(* IEC 61131-3 sources: moulding-cell-robot-interlock/plc/test/st, 1 file *)

(* ---- tb_bench.st ---- *)
(*
  TB_BENCH: self-checking test bench for the function block CELL_PLC.
  Generated by scripts/make_testbench.py from the cell model (cell/bench.py). Do not edit.

  One call is one scan of the block under test. For every scan of every case the bench applies the
  recorded input image (machine model and TP program of the repository, one PLC scan per step),
  calls its own instance of CELL_PLC and compares all outputs, the state and the fault code with
  the recorded values. A case fails at its first difference. Every case starts with a fresh instance.
  Cases: 7. Scans: 1616. Table rows (equal consecutive scans are merged): 332.
  Input bits of rowIn, from bit 0: iZA6_MouldClosed, iZA7_MouldOpenPosition, iZB2_EnableOperation, iZB3_EjectorBack, iZB4_EjectorForward, iSafetyOk, rbReqClose, rbReqEjFwd, rbReqEjBack, rbAtCut, rbPlaced, rbFault, rbAtWait, rbAreaFree, iCutClosed, iCutOpen, iNestFree, iGateClosedLocked, btnGateReq, btnReset.
  Output bits of rowExp, from bit 0: qA6_EnableMouldClosure, qB3_EnableEjectorBack, qB4_EnableEjectorForward, qB2_NoOperationWithImm, qRbImmAuto, qRbMouldOpen, qRbMouldClosed, qRbEjFwd, qRbEjBack, qRbCutDone, qRbPlaceFree, qRbCycleEnable, qRbPlaceAck, qCutClose, qConvIndex, qGateUnlock.
  rowSt = state + 16 * faultCode.
*)

FUNCTION_BLOCK TB_BENCH
VAR_INPUT
  enable : BOOL;
END_VAR
VAR_OUTPUT
  Done : BOOL;
  CasesTotal : INT;
  CasesRun : INT;
  CasesPassed : INT;
  CasesFailed : INT;
  FirstFailedCase : INT;
  FirstFailedCheck : INT;      (* scan number inside the failed case, from 1 *)
  CasePassBits : DWORD;        (* bit 0 = case 1 *)
END_VAR
VAR
  dut1 : CELL_PLC;
  dut2 : CELL_PLC;
  dut3 : CELL_PLC;
  dut4 : CELL_PLC;
  dut5 : CELL_PLC;
  dut6 : CELL_PLC;
  dut7 : CELL_PLC;
  rowIn : ARRAY [0..331] OF DWORD := [
    16#0003A02D, 16#0003A02C, 16#0003A02E, 16#0003802E, 16#000380AE, 16#000380B6, 16#00038036, 16#00038136,
    16#0003A12E, 16#0003A06E, 16#0003A06C, 16#0003A26C, 16#0003626D, 16#0003A26D, 16#0003A06D, 16#0002A06D,
    16#0002A46D, 16#0002A02D, 16#0003A02D, 16#0003A02C, 16#0003A02E, 16#0003802E, 16#000380AE, 16#000380B6,
    16#00038036, 16#00038136, 16#0003A12E, 16#0003A06E, 16#0003A06C, 16#0003A26C, 16#0003626D, 16#0003A26D,
    16#0003A06D, 16#0002A06D, 16#0002A46D, 16#0002A02D, 16#0003A02D, 16#0003A02C, 16#0003A02E, 16#0003802E,
    16#000380AE, 16#000380B6, 16#00038036, 16#00038136, 16#0003A12E, 16#0003A06E, 16#0003A06C, 16#0003A26C,
    16#0003626D, 16#0003A26D, 16#0003A06D, 16#0002A06D, 16#0002A46D, 16#0002A02D, 16#0003A02D, 16#0003A02D,
    16#0003A02C, 16#0003A02E, 16#0003802E, 16#000380AE, 16#000380B6, 16#00038036, 16#00038136, 16#0003A12E,
    16#0003A06E, 16#0003A06C, 16#0003A26C, 16#0003A26D, 16#0003A26C, 16#0003A26E, 16#0003626E, 16#0003A26E,
    16#0003A06E, 16#0002A06E, 16#0002A46E, 16#0002A02E, 16#0002A02E, 16#0003802E, 16#000380AE, 16#000380B6,
    16#00038036, 16#00038136, 16#0003A12E, 16#0003A06E, 16#0003A06C, 16#0003A26C, 16#0003A26D, 16#0003A26C,
    16#0003A26E, 16#0003626E, 16#0003A26E, 16#0003A06E, 16#0002A06E, 16#0002A46E, 16#0002A02E, 16#0002A02E,
    16#0003802E, 16#000380AE, 16#000380B6, 16#00038036, 16#00038136, 16#0003A12E, 16#0003A06E, 16#0003A06C,
    16#0003A26C, 16#0003A26D, 16#0003A02D, 16#0003A02C, 16#0003A02E, 16#0003802E, 16#000380AE, 16#000380B6,
    16#00038036, 16#00038136, 16#0003A12E, 16#0003A06E, 16#0003A06C, 16#0003A26C, 16#0003626D, 16#0003A26D,
    16#0003A06D, 16#0002A06D, 16#0002A46D, 16#0002A02D, 16#0003A02D, 16#0003A02C, 16#0003A02E, 16#0003802E,
    16#000380AE, 16#000380B6, 16#00038036, 16#00038136, 16#0003A12E, 16#0003A06E, 16#0003A06C, 16#0003826C,
    16#00038A2C, 16#0003A02D, 16#0003A02C, 16#0003A02E, 16#0003802E, 16#000380AE, 16#000380B6, 16#00038036,
    16#00038136, 16#0003A12E, 16#0003A06E, 16#0003A06C, 16#0003A26C, 16#0007626D, 16#0003626D, 16#0003A26D,
    16#0003A06D, 16#0002A06D, 16#0002A46D, 16#0002A02D, 16#0003B02D, 16#0001B02D, 16#0001B00D, 16#0001B02D,
    16#0009B02D, 16#0003B02D, 16#0003A02D, 16#0003A02C, 16#0003A02E, 16#0003802E, 16#000380AE, 16#000380B6,
    16#00038036, 16#00038136, 16#0003A12E, 16#0003A06E, 16#0003A06C, 16#0003A26C, 16#0003626D, 16#0003A26D,
    16#0003A06D, 16#0002A06D, 16#0002A46D, 16#0002A02D, 16#0003A02D, 16#0003A02C, 16#0003A02E, 16#0003802E,
    16#000380AE, 16#000380B6, 16#00038036, 16#00038136, 16#0003A12E, 16#0003A06E, 16#0003A06C, 16#0003A26C,
    16#0003626D, 16#0003A26D, 16#0003A06D, 16#0002A06D, 16#0002A46D, 16#0002A02D, 16#0003A02D, 16#0003A02D,
    16#0003A02C, 16#0003A02E, 16#0003802E, 16#000380AE, 16#000380B6, 16#00038036, 16#00038136, 16#0003A12E,
    16#0003A06E, 16#0003A06C, 16#0003A26C, 16#0003626D, 16#0003A26D, 16#0003A06D, 16#0002A06D, 16#0002A46D,
    16#0002A02D, 16#0003A02D, 16#0001A00D, 16#0003B02D, 16#000BB02D, 16#0003B02D, 16#0003A02D, 16#0003A02C,
    16#0003A02E, 16#0003802E, 16#000380AE, 16#000380B6, 16#00038036, 16#00038136, 16#0003A12E, 16#0003A06E,
    16#0003A06C, 16#0003A26C, 16#0003626D, 16#0003A26D, 16#0003A06D, 16#0002A06D, 16#0002A46D, 16#0002A02D,
    16#0003A02D, 16#0003A02C, 16#0003A02E, 16#0003802E, 16#000380AE, 16#000380B6, 16#00038036, 16#00038136,
    16#0003A12E, 16#0003A06E, 16#0003A06C, 16#0003A26C, 16#0003626D, 16#0003A26D, 16#0003A06D, 16#0002A06D,
    16#0002A46D, 16#0002A02D, 16#0003A02D, 16#0003A02D, 16#0003A02C, 16#0003A02E, 16#0003802E, 16#000380AE,
    16#000380B6, 16#00038036, 16#00038136, 16#0003A12E, 16#0003A06E, 16#0003A06C, 16#0003A26C, 16#0003626D,
    16#0003A26D, 16#0003A06D, 16#0002A06D, 16#0002A46D, 16#0002A02D, 16#0002A02C, 16#0002A02E, 16#0002802E,
    16#000280AE, 16#000280B6, 16#00028036, 16#00028136, 16#0002A12E, 16#0002A06E, 16#0002A06C, 16#0002A26C,
    16#0002626D, 16#0002A26D, 16#0002A06D, 16#0002A82D, 16#0002A82C, 16#0002A82E, 16#0003A02D, 16#0003A02C,
    16#0003A02E, 16#0003802E, 16#000380AE, 16#000380B6, 16#00038036, 16#00038136, 16#0003A12E, 16#0003A06E,
    16#0003A06C, 16#0003A26C, 16#0003626D, 16#0003A26D, 16#0003A06D, 16#0002A06D, 16#0002A46D, 16#0002A02D,
    16#0003A02D, 16#0003A02C, 16#0003A02E, 16#0003802E, 16#000380AE, 16#000380B6, 16#00038036, 16#00038136,
    16#0003A12E, 16#0003A06E, 16#0003A06C, 16#0003A26C, 16#0003626C, 16#0003A26C, 16#0003A06C, 16#0002A06C,
    16#0002A46C, 16#0002A06C, 16#0003A06C, 16#0003A82C];
  rowExp : ARRAY [0..331] OF DWORD := [
    16#00000D10, 16#00000D10, 16#00000D30, 16#00000D30, 16#00000D34, 16#00000CB4, 16#00000CB0, 16#00000CB2,
    16#00000D32, 16#00000D11, 16#00000D11, 16#00002D11, 16#00000D50, 16#00000F50, 16#00000D50, 16#00000950,
    16#00001950, 16#00005910, 16#00000D10, 16#00000D10, 16#00000D30, 16#00000D30, 16#00000D34, 16#00000CB4,
    16#00000CB0, 16#00000CB2, 16#00000D32, 16#00000D11, 16#00000D11, 16#00002D11, 16#00000D50, 16#00000F50,
    16#00000D50, 16#00000950, 16#00001950, 16#00005910, 16#00000D10, 16#00000D10, 16#00000D30, 16#00000D30,
    16#00000D34, 16#00000CB4, 16#00000CB0, 16#00000CB2, 16#00000D32, 16#00000D11, 16#00000D11, 16#00002D11,
    16#00000D50, 16#00000F50, 16#00000D50, 16#00000950, 16#00001950, 16#00005910, 16#00000D10, 16#00000D10,
    16#00000D10, 16#00000D30, 16#00000D30, 16#00000D34, 16#00000CB4, 16#00000CB0, 16#00000CB2, 16#00000D32,
    16#00000D11, 16#00000D11, 16#00002D11, 16#00002D50, 16#00002D50, 16#00002D50, 16#00000D50, 16#00000F50,
    16#00000D50, 16#00000950, 16#00001950, 16#00005910, 16#00005930, 16#00000D30, 16#00000D34, 16#00000CB4,
    16#00000CB0, 16#00000CB2, 16#00000D32, 16#00000D11, 16#00000D11, 16#00002D11, 16#00002D50, 16#00002D50,
    16#00002D50, 16#00000D50, 16#00000F50, 16#00000D50, 16#00000950, 16#00001950, 16#00005910, 16#00005930,
    16#00000D30, 16#00000D34, 16#00000CB4, 16#00000CB0, 16#00000CB2, 16#00000D32, 16#00000D11, 16#00000D11,
    16#00002D11, 16#00002D50, 16#00000D10, 16#00000D10, 16#00000D30, 16#00000D30, 16#00000D34, 16#00000CB4,
    16#00000CB0, 16#00000CB2, 16#00000D32, 16#00000D11, 16#00000D11, 16#00002D11, 16#00000D50, 16#00000F50,
    16#00000D50, 16#00000950, 16#00001950, 16#00005910, 16#00000D10, 16#00000D10, 16#00000D30, 16#00000D30,
    16#00000D34, 16#00000CB4, 16#00000CB0, 16#00000CB2, 16#00000D32, 16#00000D11, 16#00000D11, 16#00000500,
    16#00000500, 16#00000D10, 16#00000D10, 16#00000D30, 16#00000D30, 16#00000D34, 16#00000CB4, 16#00000CB0,
    16#00000CB2, 16#00000D32, 16#00000D11, 16#00000D11, 16#00002D11, 16#00000550, 16#00000550, 16#00000750,
    16#00000550, 16#00000150, 16#00001150, 16#00005110, 16#00008500, 16#00008500, 16#00008500, 16#00008500,
    16#00000500, 16#00000D10, 16#00000D10, 16#00000D10, 16#00000D30, 16#00000D30, 16#00000D34, 16#00000CB4,
    16#00000CB0, 16#00000CB2, 16#00000D32, 16#00000D11, 16#00000D11, 16#00002D11, 16#00000D50, 16#00000F50,
    16#00000D50, 16#00000950, 16#00001950, 16#00005910, 16#00000D10, 16#00000D10, 16#00000D30, 16#00000D30,
    16#00000D34, 16#00000CB4, 16#00000CB0, 16#00000CB2, 16#00000D32, 16#00000D11, 16#00000D11, 16#00002D11,
    16#00000D50, 16#00000F50, 16#00000D50, 16#00000950, 16#00001950, 16#00005910, 16#00000D10, 16#00000D10,
    16#00000D10, 16#00000D30, 16#00000D30, 16#00000D34, 16#00000CB4, 16#00000CB0, 16#00000CB2, 16#00000D32,
    16#00000D11, 16#00000D11, 16#00002D11, 16#00000D50, 16#00000F50, 16#00000D50, 16#00000950, 16#00001950,
    16#00005910, 16#00000D10, 16#00000500, 16#00000500, 16#00000500, 16#00000D10, 16#00000D10, 16#00000D10,
    16#00000D30, 16#00000D30, 16#00000D34, 16#00000CB4, 16#00000CB0, 16#00000CB2, 16#00000D32, 16#00000D11,
    16#00000D11, 16#00002D11, 16#00000D50, 16#00000F50, 16#00000D50, 16#00000950, 16#00001950, 16#00005910,
    16#00000D10, 16#00000D10, 16#00000D30, 16#00000D30, 16#00000D34, 16#00000CB4, 16#00000CB0, 16#00000CB2,
    16#00000D32, 16#00000D11, 16#00000D11, 16#00002D11, 16#00000D50, 16#00000F50, 16#00000D50, 16#00000950,
    16#00001950, 16#00005910, 16#00000D10, 16#00000D10, 16#00000D10, 16#00000D30, 16#00000D30, 16#00000D34,
    16#00000CB4, 16#00000CB0, 16#00000CB2, 16#00000D32, 16#00000D11, 16#00000D11, 16#00002D11, 16#00000D50,
    16#00000F50, 16#00000D50, 16#00000950, 16#00001950, 16#00005910, 16#00005910, 16#00005930, 16#00005930,
    16#00005934, 16#000058B4, 16#000058B0, 16#000058B2, 16#00005932, 16#00005911, 16#00005911, 16#00007911,
    16#00005950, 16#00005B50, 16#00005950, 16#00001140, 16#00001140, 16#00001140, 16#00000D10, 16#00000D10,
    16#00000D30, 16#00000D30, 16#00000D34, 16#00000CB4, 16#00000CB0, 16#00000CB2, 16#00000D32, 16#00000D11,
    16#00000D11, 16#00002D11, 16#00000D50, 16#00000F50, 16#00000D50, 16#00000950, 16#00001950, 16#00005910,
    16#00000D10, 16#00000D10, 16#00000D30, 16#00000D30, 16#00000D34, 16#00000CB4, 16#00000CB0, 16#00000CB2,
    16#00000D32, 16#00000D11, 16#00000D11, 16#00002D11, 16#00000D11, 16#00000F11, 16#00000D11, 16#00000911,
    16#00001911, 16#00005911, 16#00000500, 16#00000500];
  rowSt : ARRAY [0..331] OF INT := [
    1, 1, 2, 3, 3, 3, 3, 3, 3, 4, 4, 4, 1, 1, 1, 1, 1, 1, 1, 1,
    2, 3, 3, 3, 3, 3, 3, 4, 4, 4, 1, 1, 1, 1, 1, 1, 1, 1, 2, 3,
    3, 3, 3, 3, 3, 4, 4, 4, 1, 1, 1, 1, 1, 1, 1, 1, 1, 2, 3, 3,
    3, 3, 3, 3, 4, 4, 4, 1, 1, 1, 1, 1, 1, 1, 1, 1, 2, 3, 3, 3,
    3, 3, 3, 4, 4, 4, 1, 1, 1, 1, 1, 1, 1, 1, 1, 2, 3, 3, 3, 3,
    3, 3, 4, 4, 4, 1, 1, 1, 2, 3, 3, 3, 3, 3, 3, 4, 4, 4, 1, 1,
    1, 1, 1, 1, 1, 1, 2, 3, 3, 3, 3, 3, 3, 4, 4, 89, 89, 1, 1, 2,
    3, 3, 3, 3, 3, 3, 4, 4, 4, 1, 1, 1, 1, 1, 1, 1, 5, 5, 5, 5,
    5, 1, 1, 1, 2, 3, 3, 3, 3, 3, 3, 4, 4, 4, 1, 1, 1, 1, 1, 1,
    1, 1, 2, 3, 3, 3, 3, 3, 3, 4, 4, 4, 1, 1, 1, 1, 1, 1, 1, 1,
    1, 2, 3, 3, 3, 3, 3, 3, 4, 4, 4, 1, 1, 1, 1, 1, 1, 1, 25, 25,
    16, 1, 1, 1, 2, 3, 3, 3, 3, 3, 3, 4, 4, 4, 1, 1, 1, 1, 1, 1,
    1, 1, 2, 3, 3, 3, 3, 3, 3, 4, 4, 4, 1, 1, 1, 1, 1, 1, 1, 1,
    1, 2, 3, 3, 3, 3, 3, 3, 4, 4, 4, 1, 1, 1, 1, 1, 1, 1, 2, 3,
    3, 3, 3, 3, 3, 4, 4, 4, 1, 1, 1, 41, 41, 41, 1, 1, 2, 3, 3, 3,
    3, 3, 3, 4, 4, 4, 1, 1, 1, 1, 1, 1, 1, 1, 2, 3, 3, 3, 3, 3,
    3, 4, 4, 4, 4, 4, 4, 4, 4, 4, 105, 105];
  rowRep : ARRAY [0..331] OF INT := [
    45, 4, 1, 6, 3, 1, 3, 3, 1, 1, 2, 3, 3, 1, 8, 3, 1, 4, 25, 4,
    1, 6, 3, 1, 3, 3, 1, 1, 2, 3, 3, 1, 8, 3, 1, 4, 25, 4, 1, 6,
    3, 1, 3, 3, 1, 1, 2, 3, 3, 1, 8, 3, 1, 4, 7, 45, 4, 1, 6, 3,
    1, 3, 3, 1, 1, 2, 3, 45, 4, 9, 3, 1, 8, 3, 1, 1, 3, 6, 3, 1,
    3, 3, 1, 1, 2, 3, 45, 4, 9, 3, 1, 8, 3, 1, 1, 3, 6, 3, 1, 3,
    3, 1, 1, 2, 3, 7, 45, 4, 1, 6, 3, 1, 3, 3, 1, 1, 2, 3, 3, 1,
    8, 3, 1, 4, 25, 4, 1, 6, 3, 1, 3, 3, 1, 1, 2, 40, 7, 45, 4, 1,
    6, 3, 1, 3, 3, 1, 1, 2, 3, 1, 2, 1, 8, 3, 1, 4, 1, 3, 6, 3,
    1, 1, 10, 4, 1, 6, 3, 1, 3, 3, 1, 1, 2, 3, 3, 1, 8, 3, 1, 4,
    25, 4, 1, 6, 3, 1, 3, 3, 1, 1, 2, 3, 3, 1, 8, 3, 1, 4, 7, 45,
    4, 1, 6, 3, 1, 3, 3, 1, 1, 2, 3, 3, 1, 8, 3, 1, 4, 3, 6, 4,
    1, 1, 10, 4, 1, 6, 3, 1, 3, 3, 1, 1, 2, 3, 3, 1, 8, 3, 1, 4,
    25, 4, 1, 6, 3, 1, 3, 3, 1, 1, 2, 3, 3, 1, 8, 3, 1, 4, 7, 45,
    4, 1, 6, 3, 1, 3, 3, 1, 1, 2, 3, 3, 1, 8, 3, 1, 29, 4, 1, 6,
    3, 1, 3, 3, 1, 1, 2, 3, 3, 1, 40, 1, 4, 2, 45, 4, 1, 6, 3, 1,
    3, 3, 1, 1, 2, 3, 3, 1, 8, 3, 1, 4, 25, 4, 1, 6, 3, 1, 3, 3,
    1, 1, 2, 3, 3, 1, 8, 3, 1, 4, 36, 7];
  caseFirst : ARRAY [1..7] OF INT := [0, 55, 106, 137, 199, 259, 294];
  caseLast : ARRAY [1..7] OF INT := [54, 105, 136, 198, 258, 293, 331];
  caseMask : ARRAY [1..7] OF DWORD := [16#00000001, 16#00000002, 16#00000004, 16#00000008, 16#00000010, 16#00000020, 16#00000040];
  c : INT := 1;
  r : INT;
  k : INT;
  check : INT;
  started : BOOL;
  finished : BOOL;
  caseEnd : BOOL;
  nRun : INT;
  nPass : INT;
  nFail : INT;
  ffCase : INT;
  ffCheck : INT;
  passBits : DWORD;
  w : DWORD;
  got : DWORD;
  gotSt : INT;
  oState : INT;
  oFault : INT;
  i0 : BOOL;
  i1 : BOOL;
  i2 : BOOL;
  i3 : BOOL;
  i4 : BOOL;
  i5 : BOOL;
  i6 : BOOL;
  i7 : BOOL;
  i8 : BOOL;
  i9 : BOOL;
  i10 : BOOL;
  i11 : BOOL;
  i12 : BOOL;
  i13 : BOOL;
  i14 : BOOL;
  i15 : BOOL;
  i16 : BOOL;
  i17 : BOOL;
  i18 : BOOL;
  i19 : BOOL;
  o0 : BOOL;
  o1 : BOOL;
  o2 : BOOL;
  o3 : BOOL;
  o4 : BOOL;
  o5 : BOOL;
  o6 : BOOL;
  o7 : BOOL;
  o8 : BOOL;
  o9 : BOOL;
  o10 : BOOL;
  o11 : BOOL;
  o12 : BOOL;
  o13 : BOOL;
  o14 : BOOL;
  o15 : BOOL;
END_VAR

  IF enable AND NOT finished THEN
    IF NOT started THEN
      started := TRUE;
      r := caseFirst[c];
      k := 0;
      check := 0;
    END_IF;

    (* input image of this scan *)
    w := rowIn[r];
    i0 := (w AND DWORD#1) <> DWORD#0;
    i1 := (w AND DWORD#2) <> DWORD#0;
    i2 := (w AND DWORD#4) <> DWORD#0;
    i3 := (w AND DWORD#8) <> DWORD#0;
    i4 := (w AND DWORD#16) <> DWORD#0;
    i5 := (w AND DWORD#32) <> DWORD#0;
    i6 := (w AND DWORD#64) <> DWORD#0;
    i7 := (w AND DWORD#128) <> DWORD#0;
    i8 := (w AND DWORD#256) <> DWORD#0;
    i9 := (w AND DWORD#512) <> DWORD#0;
    i10 := (w AND DWORD#1024) <> DWORD#0;
    i11 := (w AND DWORD#2048) <> DWORD#0;
    i12 := (w AND DWORD#4096) <> DWORD#0;
    i13 := (w AND DWORD#8192) <> DWORD#0;
    i14 := (w AND DWORD#16384) <> DWORD#0;
    i15 := (w AND DWORD#32768) <> DWORD#0;
    i16 := (w AND DWORD#65536) <> DWORD#0;
    i17 := (w AND DWORD#131072) <> DWORD#0;
    i18 := (w AND DWORD#262144) <> DWORD#0;
    i19 := (w AND DWORD#524288) <> DWORD#0;

    (* one scan of the block under test *)
    CASE c OF
      1:
        dut1(iZA6_MouldClosed := i0, iZA7_MouldOpenPosition := i1, iZB2_EnableOperation := i2, iZB3_EjectorBack := i3, iZB4_EjectorForward := i4, iSafetyOk := i5, rbReqClose := i6, rbReqEjFwd := i7, rbReqEjBack := i8, rbAtCut := i9, rbPlaced := i10, rbFault := i11, rbAtWait := i12, rbAreaFree := i13, iCutClosed := i14, iCutOpen := i15, iNestFree := i16, iGateClosedLocked := i17, btnGateReq := i18, btnReset := i19, cfgCloseTmoScans := 25);
        o0 := dut1.qA6_EnableMouldClosure;
        o1 := dut1.qB3_EnableEjectorBack;
        o2 := dut1.qB4_EnableEjectorForward;
        o3 := dut1.qB2_NoOperationWithImm;
        o4 := dut1.qRbImmAuto;
        o5 := dut1.qRbMouldOpen;
        o6 := dut1.qRbMouldClosed;
        o7 := dut1.qRbEjFwd;
        o8 := dut1.qRbEjBack;
        o9 := dut1.qRbCutDone;
        o10 := dut1.qRbPlaceFree;
        o11 := dut1.qRbCycleEnable;
        o12 := dut1.qRbPlaceAck;
        o13 := dut1.qCutClose;
        o14 := dut1.qConvIndex;
        o15 := dut1.qGateUnlock;
        oState := dut1.state;
        oFault := dut1.faultCode;
      2:
        dut2(iZA6_MouldClosed := i0, iZA7_MouldOpenPosition := i1, iZB2_EnableOperation := i2, iZB3_EjectorBack := i3, iZB4_EjectorForward := i4, iSafetyOk := i5, rbReqClose := i6, rbReqEjFwd := i7, rbReqEjBack := i8, rbAtCut := i9, rbPlaced := i10, rbFault := i11, rbAtWait := i12, rbAreaFree := i13, iCutClosed := i14, iCutOpen := i15, iNestFree := i16, iGateClosedLocked := i17, btnGateReq := i18, btnReset := i19, cfgCloseTmoScans := 25);
        o0 := dut2.qA6_EnableMouldClosure;
        o1 := dut2.qB3_EnableEjectorBack;
        o2 := dut2.qB4_EnableEjectorForward;
        o3 := dut2.qB2_NoOperationWithImm;
        o4 := dut2.qRbImmAuto;
        o5 := dut2.qRbMouldOpen;
        o6 := dut2.qRbMouldClosed;
        o7 := dut2.qRbEjFwd;
        o8 := dut2.qRbEjBack;
        o9 := dut2.qRbCutDone;
        o10 := dut2.qRbPlaceFree;
        o11 := dut2.qRbCycleEnable;
        o12 := dut2.qRbPlaceAck;
        o13 := dut2.qCutClose;
        o14 := dut2.qConvIndex;
        o15 := dut2.qGateUnlock;
        oState := dut2.state;
        oFault := dut2.faultCode;
      3:
        dut3(iZA6_MouldClosed := i0, iZA7_MouldOpenPosition := i1, iZB2_EnableOperation := i2, iZB3_EjectorBack := i3, iZB4_EjectorForward := i4, iSafetyOk := i5, rbReqClose := i6, rbReqEjFwd := i7, rbReqEjBack := i8, rbAtCut := i9, rbPlaced := i10, rbFault := i11, rbAtWait := i12, rbAreaFree := i13, iCutClosed := i14, iCutOpen := i15, iNestFree := i16, iGateClosedLocked := i17, btnGateReq := i18, btnReset := i19, cfgCloseTmoScans := 25);
        o0 := dut3.qA6_EnableMouldClosure;
        o1 := dut3.qB3_EnableEjectorBack;
        o2 := dut3.qB4_EnableEjectorForward;
        o3 := dut3.qB2_NoOperationWithImm;
        o4 := dut3.qRbImmAuto;
        o5 := dut3.qRbMouldOpen;
        o6 := dut3.qRbMouldClosed;
        o7 := dut3.qRbEjFwd;
        o8 := dut3.qRbEjBack;
        o9 := dut3.qRbCutDone;
        o10 := dut3.qRbPlaceFree;
        o11 := dut3.qRbCycleEnable;
        o12 := dut3.qRbPlaceAck;
        o13 := dut3.qCutClose;
        o14 := dut3.qConvIndex;
        o15 := dut3.qGateUnlock;
        oState := dut3.state;
        oFault := dut3.faultCode;
      4:
        dut4(iZA6_MouldClosed := i0, iZA7_MouldOpenPosition := i1, iZB2_EnableOperation := i2, iZB3_EjectorBack := i3, iZB4_EjectorForward := i4, iSafetyOk := i5, rbReqClose := i6, rbReqEjFwd := i7, rbReqEjBack := i8, rbAtCut := i9, rbPlaced := i10, rbFault := i11, rbAtWait := i12, rbAreaFree := i13, iCutClosed := i14, iCutOpen := i15, iNestFree := i16, iGateClosedLocked := i17, btnGateReq := i18, btnReset := i19, cfgCloseTmoScans := 25);
        o0 := dut4.qA6_EnableMouldClosure;
        o1 := dut4.qB3_EnableEjectorBack;
        o2 := dut4.qB4_EnableEjectorForward;
        o3 := dut4.qB2_NoOperationWithImm;
        o4 := dut4.qRbImmAuto;
        o5 := dut4.qRbMouldOpen;
        o6 := dut4.qRbMouldClosed;
        o7 := dut4.qRbEjFwd;
        o8 := dut4.qRbEjBack;
        o9 := dut4.qRbCutDone;
        o10 := dut4.qRbPlaceFree;
        o11 := dut4.qRbCycleEnable;
        o12 := dut4.qRbPlaceAck;
        o13 := dut4.qCutClose;
        o14 := dut4.qConvIndex;
        o15 := dut4.qGateUnlock;
        oState := dut4.state;
        oFault := dut4.faultCode;
      5:
        dut5(iZA6_MouldClosed := i0, iZA7_MouldOpenPosition := i1, iZB2_EnableOperation := i2, iZB3_EjectorBack := i3, iZB4_EjectorForward := i4, iSafetyOk := i5, rbReqClose := i6, rbReqEjFwd := i7, rbReqEjBack := i8, rbAtCut := i9, rbPlaced := i10, rbFault := i11, rbAtWait := i12, rbAreaFree := i13, iCutClosed := i14, iCutOpen := i15, iNestFree := i16, iGateClosedLocked := i17, btnGateReq := i18, btnReset := i19, cfgCloseTmoScans := 25);
        o0 := dut5.qA6_EnableMouldClosure;
        o1 := dut5.qB3_EnableEjectorBack;
        o2 := dut5.qB4_EnableEjectorForward;
        o3 := dut5.qB2_NoOperationWithImm;
        o4 := dut5.qRbImmAuto;
        o5 := dut5.qRbMouldOpen;
        o6 := dut5.qRbMouldClosed;
        o7 := dut5.qRbEjFwd;
        o8 := dut5.qRbEjBack;
        o9 := dut5.qRbCutDone;
        o10 := dut5.qRbPlaceFree;
        o11 := dut5.qRbCycleEnable;
        o12 := dut5.qRbPlaceAck;
        o13 := dut5.qCutClose;
        o14 := dut5.qConvIndex;
        o15 := dut5.qGateUnlock;
        oState := dut5.state;
        oFault := dut5.faultCode;
      6:
        dut6(iZA6_MouldClosed := i0, iZA7_MouldOpenPosition := i1, iZB2_EnableOperation := i2, iZB3_EjectorBack := i3, iZB4_EjectorForward := i4, iSafetyOk := i5, rbReqClose := i6, rbReqEjFwd := i7, rbReqEjBack := i8, rbAtCut := i9, rbPlaced := i10, rbFault := i11, rbAtWait := i12, rbAreaFree := i13, iCutClosed := i14, iCutOpen := i15, iNestFree := i16, iGateClosedLocked := i17, btnGateReq := i18, btnReset := i19, cfgCloseTmoScans := 25);
        o0 := dut6.qA6_EnableMouldClosure;
        o1 := dut6.qB3_EnableEjectorBack;
        o2 := dut6.qB4_EnableEjectorForward;
        o3 := dut6.qB2_NoOperationWithImm;
        o4 := dut6.qRbImmAuto;
        o5 := dut6.qRbMouldOpen;
        o6 := dut6.qRbMouldClosed;
        o7 := dut6.qRbEjFwd;
        o8 := dut6.qRbEjBack;
        o9 := dut6.qRbCutDone;
        o10 := dut6.qRbPlaceFree;
        o11 := dut6.qRbCycleEnable;
        o12 := dut6.qRbPlaceAck;
        o13 := dut6.qCutClose;
        o14 := dut6.qConvIndex;
        o15 := dut6.qGateUnlock;
        oState := dut6.state;
        oFault := dut6.faultCode;
      7:
        dut7(iZA6_MouldClosed := i0, iZA7_MouldOpenPosition := i1, iZB2_EnableOperation := i2, iZB3_EjectorBack := i3, iZB4_EjectorForward := i4, iSafetyOk := i5, rbReqClose := i6, rbReqEjFwd := i7, rbReqEjBack := i8, rbAtCut := i9, rbPlaced := i10, rbFault := i11, rbAtWait := i12, rbAreaFree := i13, iCutClosed := i14, iCutOpen := i15, iNestFree := i16, iGateClosedLocked := i17, btnGateReq := i18, btnReset := i19, cfgCloseTmoScans := 25);
        o0 := dut7.qA6_EnableMouldClosure;
        o1 := dut7.qB3_EnableEjectorBack;
        o2 := dut7.qB4_EnableEjectorForward;
        o3 := dut7.qB2_NoOperationWithImm;
        o4 := dut7.qRbImmAuto;
        o5 := dut7.qRbMouldOpen;
        o6 := dut7.qRbMouldClosed;
        o7 := dut7.qRbEjFwd;
        o8 := dut7.qRbEjBack;
        o9 := dut7.qRbCutDone;
        o10 := dut7.qRbPlaceFree;
        o11 := dut7.qRbCycleEnable;
        o12 := dut7.qRbPlaceAck;
        o13 := dut7.qCutClose;
        o14 := dut7.qConvIndex;
        o15 := dut7.qGateUnlock;
        oState := dut7.state;
        oFault := dut7.faultCode;
    END_CASE;

    (* output image *)
    got := DWORD#0;
    IF o0 THEN
      got := got OR DWORD#1;
    END_IF;
    IF o1 THEN
      got := got OR DWORD#2;
    END_IF;
    IF o2 THEN
      got := got OR DWORD#4;
    END_IF;
    IF o3 THEN
      got := got OR DWORD#8;
    END_IF;
    IF o4 THEN
      got := got OR DWORD#16;
    END_IF;
    IF o5 THEN
      got := got OR DWORD#32;
    END_IF;
    IF o6 THEN
      got := got OR DWORD#64;
    END_IF;
    IF o7 THEN
      got := got OR DWORD#128;
    END_IF;
    IF o8 THEN
      got := got OR DWORD#256;
    END_IF;
    IF o9 THEN
      got := got OR DWORD#512;
    END_IF;
    IF o10 THEN
      got := got OR DWORD#1024;
    END_IF;
    IF o11 THEN
      got := got OR DWORD#2048;
    END_IF;
    IF o12 THEN
      got := got OR DWORD#4096;
    END_IF;
    IF o13 THEN
      got := got OR DWORD#8192;
    END_IF;
    IF o14 THEN
      got := got OR DWORD#16384;
    END_IF;
    IF o15 THEN
      got := got OR DWORD#32768;
    END_IF;
    gotSt := oState + 16 * oFault;

    (* compare, then step through the table *)
    check := check + 1;
    k := k + 1;
    caseEnd := FALSE;
    IF got <> rowExp[r] OR gotSt <> rowSt[r] THEN
      nFail := nFail + 1;
      IF ffCase = 0 THEN
        ffCase := c;
        ffCheck := check;
      END_IF;
      caseEnd := TRUE;
    ELSIF k >= rowRep[r] THEN
      k := 0;
      IF r >= caseLast[c] THEN
        nPass := nPass + 1;
        passBits := passBits OR caseMask[c];
        caseEnd := TRUE;
      ELSE
        r := r + 1;
      END_IF;
    END_IF;
    IF caseEnd THEN
      nRun := nRun + 1;
      started := FALSE;
      IF c >= 7 THEN
        finished := TRUE;
      ELSE
        c := c + 1;
      END_IF;
    END_IF;
  END_IF;

  (* outputs are written once and never read back; the result is held after the last case *)
  Done := finished;
  CasesTotal := 7;
  CasesRun := nRun;
  CasesPassed := nPass;
  CasesFailed := nFail;
  FirstFailedCase := ffCase;
  FirstFailedCheck := ffCheck;
  CasePassBits := passBits;
END_FUNCTION_BLOCK
